(* IEC 61131-3 sources: s7-to-codesys/tests/POUs/S7Compat/FB_S7FTrig_Test, 3 files *)

(* ---- FallingEdgeOnce.method.decl.st ---- *)
// TRUE -> FALSE: Q = TRUE ровно на одном вызове.
METHOD PRIVATE FallingEdgeOnce
VAR
    fbDut : FB_S7FTrig;     // проверяемый детектор (новый экземпляр на каждый вызов метода)
END_VAR

(* ---- NoEdgeOnFirstCallWithClkFalse.method.decl.st ---- *)
// семантика S7: на первом вызове с CLK = FALSE спада нет.
METHOD PRIVATE NoEdgeOnFirstCallWithClkFalse
VAR
    fbDut : FB_S7FTrig;     // проверяемый детектор (новый экземпляр на каждый вызов метода)
END_VAR

(* ---- StandardFTrigMatchesS7.method.decl.st ---- *)
// Характеризация платформы: F_TRIG библиотеки Standard CODESYS на тех же входах, что и FB_S7FTrig
// (семантика S7): на первом вызове с CLK = FALSE спада нет, спад TRUE -> FALSE — ровно на одном вызове.
// Если тест упадёт на другой версии Standard, корпус собирают с --f-trig s7compat (docs/MAPPING.md, fb.f_trig).
METHOD PRIVATE StandardFTrigMatchesS7
VAR
    fbStandard : F_TRIG;    // F_TRIG библиотеки Standard (новый экземпляр на каждый вызов метода)
    fbCompat : FB_S7FTrig;  // эталон семантики S7
END_VAR
